(* PLC project Unnamed, Unknown Unnamed 1 *)
(* stored: creationDateTime 2025-10-06T15:49:55, modificationDateTime 2025-10-07T22:20:17 *)

PROGRAM program0
  VAR
    valveA AT %QX0.1 : BOOL;
    valveB AT %QX0.2 : BOOL;
    valveC AT %QX0.3 : BOOL;
    alarm AT %QX0.6 : BOOL;
    indicator AT %QX0.0 : BOOL;
    start AT %IX0.0 : BOOL;
    stop AT %IX0.1 : BOOL;
  END_VAR
  VAR_EXTERNAL
    valveAext : BOOL;
    valveBext : BOOL;
    valveCext : BOOL;
  END_VAR
  VAR
    mixer AT %QX0.4 : BOOL;
    heater AT %QX0.5 : BOOL;
  END_VAR
  VAR_EXTERNAL
    heaterExt : BOOL;
    level : INT;
  END_VAR
  VAR
    level0 AT %MW0 : INT;
  END_VAR
  VAR_EXTERNAL
    temp : INT;
  END_VAR
  VAR
    temp0 : INT;
  END_VAR
  VAR
    tempSet AT %IW0 : INT;
    tempSet0 AT %IW1 : INT;
  END_VAR
  VAR
    TOF0 : TOF;
    TP1 : TP;
    CTU0 : CTU;
  END_VAR
  VAR  (* added by the conversion: wires and edge detectors of the diagram *)
    R_TRIG1 : R_TRIG;
    R_TRIG2 : R_TRIG;
    R_TRIG3 : R_TRIG;
    F_TRIG4 : F_TRIG;
    F_TRIG5 : F_TRIG;
    F_TRIG6 : F_TRIG;
    F_TRIG7 : F_TRIG;
    F_TRIG8 : F_TRIG;
    R_TRIG9 : R_TRIG;
  END_VAR

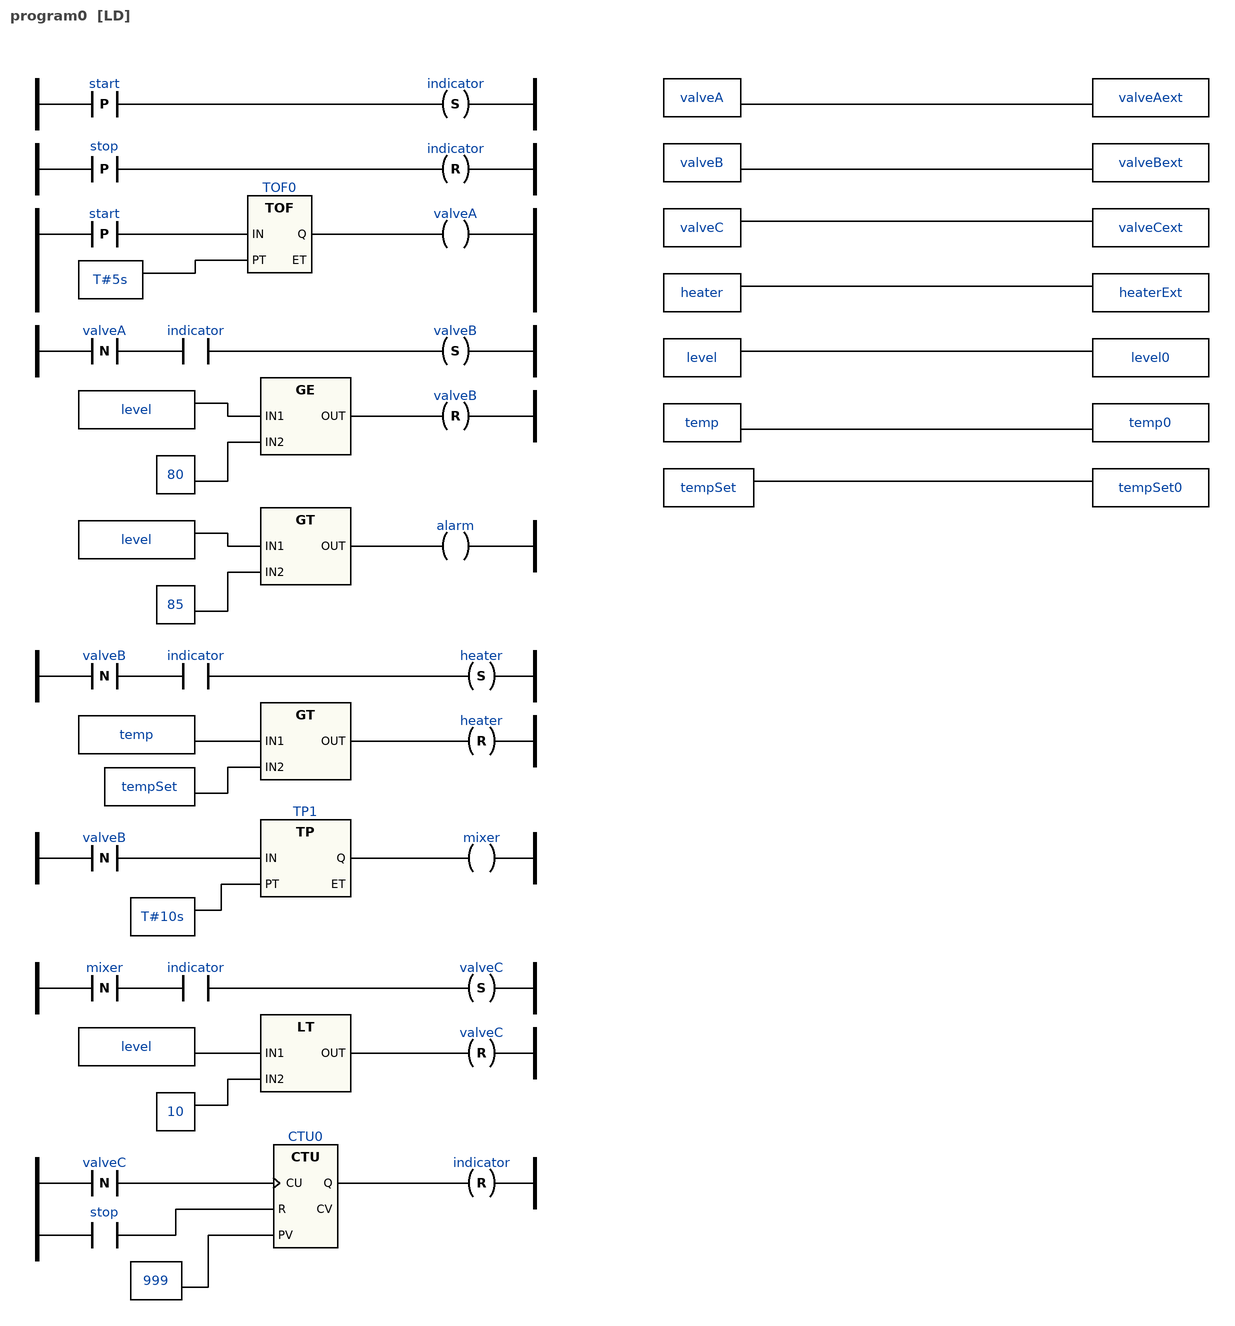
(* LD diagram, written out as Structured Text *)
R_TRIG1(CLK := start);
IF R_TRIG1.Q THEN indicator := TRUE; END_IF;
valveAext := valveA;
R_TRIG2(CLK := stop);
IF R_TRIG2.Q THEN indicator := FALSE; END_IF;
R_TRIG3(CLK := start);
TOF0(IN := R_TRIG3.Q, PT := T#5s);
valveA := TOF0.Q;
F_TRIG4(CLK := valveA);
IF F_TRIG4.Q AND indicator THEN valveB := TRUE; END_IF;
IF level >= 80 THEN valveB := FALSE; END_IF;
alarm := level > 85;
valveBext := valveB;
F_TRIG5(CLK := valveB);
IF F_TRIG5.Q AND indicator THEN heater := TRUE; END_IF;
IF temp > tempSet THEN heater := FALSE; END_IF;
heaterExt := heater;
F_TRIG6(CLK := valveB);
TP1(IN := F_TRIG6.Q, PT := T#10s);
mixer := TP1.Q;
F_TRIG7(CLK := mixer);
IF F_TRIG7.Q AND indicator THEN valveC := TRUE; END_IF;
IF level < 10 THEN valveC := FALSE; END_IF;
valveCext := valveC;
F_TRIG8(CLK := valveC);
R_TRIG9(CLK := F_TRIG8.Q);
CTU0(CU := R_TRIG9.Q, R := stop, PV := 999);
IF CTU0.Q THEN indicator := FALSE; END_IF;
level0 := level;
temp0 := temp;
tempSet0 := tempSet;
END_PROGRAM

CONFIGURATION Config0
  RESOURCE Res0 ON PLC
    TASK task0(INTERVAL := T#100ms, PRIORITY := 0);
    PROGRAM instance0 WITH task0 : program0;
  END_RESOURCE
END_CONFIGURATION
